TYPE ST_AxisCalibrationRecord :
STRUCT
SchemaVersion : UDINT;
AxisKey : STRING(63);
BaselineVersion : UDINT;
ScaleFingerprint : STRING(63);
Scale : LREAL;
EncoderOffset : LREAL;
EncoderInverse : BOOL;
Modulo : LREAL;
Offset : LREAL;
Revision : UDINT;
Integrity : DWORD;
END_STRUCT
END_TYPE

(* stored: Version 1.1.0.1, ProductVersion 3.1.4026.20
   DUT ST_AxisCalibrationRecord: Id {7f4ede88-b60a-5567-b856-0c5b4b99743e} *)
